(* IEC 61131-3 sources: WenQuest/textbook/plc/ch04/code, 3 files *)

(* ---- p4_3_1.st ---- *)
(* 程序 4.3.1  计件，外加一段“别的工作”：FOR 循环执行 n 次，用来模拟程序变长（数据记录、通信处理……） *)
PROGRAM Main
  VAR
    cnt : CTU;            (* 工件计数 *)
    n : DINT := 1000;     (* “别的工作”的循环次数：改它，看扫描时间怎样变 *)
    i : DINT;
    work : DINT;
  END_VAR
  cnt(CU := B1_Part, R := S1_Reset, PV := 30000);
  FOR i := 1 TO n DO
    work := work + 1;
  END_FOR;
  H1_Count := B1_Part;
END_PROGRAM

(* ---- p4_6_1.st ---- *)
(* 程序 4.6.1  扫描带来的三件“怪事”：一拍延迟、双线圈、程序顺序决定结果 *)
PROGRAM Main
  (* 1. 一拍延迟：H2 用的是 H1 上一次扫描的值 *)
  H2_Late := H1_Copy;
  H1_Copy := S1_In;

  (* 2. 双线圈：Y1 被写了两次，只有后一次起作用 *)
  Y1_Out := S1_In;
  Y1_Out := S2_In;

  (* 3. 顺序：先算 H3_First，再用它，就没有延迟 *)
  H3_First := S1_In;
  H4_Same := H3_First;
END_PROGRAM

(* ---- p4_7_1.st ---- *)
(* 程序 4.7.1  计件：普通输入 + 计数器（原程序）与读高速计数器（改后）并排 *)
PROGRAM Main
  VAR
    cnt : CTU;                 (* 原程序：对 B1_Part 的上升沿计数，每次扫描看一次 *)
    base : DINT;               (* 改后：清零时记下高速计数器的读数 *)
    countHsc : DINT;          (* 改后：本班的件数 *)
    n : DINT := 5000;          (* 其余程序，用一个循环代替，使扫描时间约 10 ms *)
    i : DINT;
    work : DINT;
  END_VAR
  cnt(CU := B1_Part, R := S1_Reset, PV := 30000);

  IF S1_Reset THEN
    base := HSC1_CV;
  END_IF;
  countHsc := HSC1_CV - base;

  FOR i := 1 TO n DO
    work := work + 1;
  END_FOR;
  H1_Count := B1_Part;
END_PROGRAM
